# EPICS substitutions: b-55B2VNC/src/main/epics/PCF0CoreApp/Db/Ni5763_NDS_DAN_Plugin.substitutions
file "nds3_StateMachine.template" {
pattern
{
    BOARDTYPE,
    BOARDTYPEIDX,
    CBS1,
    CBS2,
    STATEMACHINE_NAME
}
{
    "NDSDAN",
    "0",
    "D1",
    "I2",
    "StateMachine"
}
}
